Staubli VAL3: main.pgx

program main()
begin
  close(tCurrentTool)
  pPointRx.config.shoulder = lefty
  pPointRx.config.elbow = epositive
  pPointRx.config.wrist = wpositive
  pPointRx2.config.shoulder = lefty
  pPointRx2.config.elbow = epositive
  pPointRx2.config.wrist = wpositive
  mCurrentSpeed.tvel = 100.00
  mCurrentSpeed.blend = joint
  mCurrentSpeed.reach = 0.010
  mCurrentSpeed.leave = 0.010
  call MoveJoint(20.00000,-10.00000,20.00000,0.00000,30.00000,0.00000)
  call MoveJoint(0.00000,-10.00000,20.00000,0.00000,30.00000,0.00000)
  call MoveJoint(20.00000,-10.00000,20.00000,0.00000,30.00000,0.00000)
  call MoveJoint(0.00000,-10.00000,20.00000,0.00000,30.00000,0.00000)
  call MoveJoint(20.00000,-10.00000,20.00000,0.00000,30.00000,0.00000)
  call MoveJoint(0.00000,-10.00000,20.00000,0.00000,30.00000,0.00000)

end
